(* IEC 61131-3 sources: machine-design-framework/examples/pick-glue-place/plc/generated, 2 files *)

(* ---- GVL_Cycle.st ---- *)
(* GENERATED from cycle.yaml - DO NOT EDIT. source-hash: bd31026db604f3bd *)
(* Commanded angles (deg). Effective timing = commanded + device delay; see GLUE-BEAD/PROD-* checks. *)
VAR_GLOBAL CONSTANT
    VACUUM_ON  : REAL := 10.0000;
    VACUUM_OFF : REAL := 222.0000;
    GLUE_GUN_ON  : REAL := 128.6400;
    GLUE_GUN_OFF : REAL := 130.4000;
    VAC_OK_CHECK : REAL := 26.0000;
    DOUBLE_SHEET_CHECK : REAL := 75.0000;
    HOST_BOOK_CHECK : REAL := 5.0000;
    HOST_SPINE_CHECK : REAL := 140.0000;
    BEAD_OK_CHECK : REAL := 148.0000;
    X_TRANSFER_OFFSET_MIN : REAL := 0.0000;   (* per-cycle offset range, mm *)
    X_TRANSFER_OFFSET_MAX : REAL := 15.0000;
    PARK_ANGLE : REAL := 355.0000;
END_VAR

(* ---- GVL_IO.st ---- *)
(* GENERATED from io_list.yaml - DO NOT EDIT. source-hash: db4df5e0d0977f7a *)
VAR_GLOBAL
    rAngle : REAL;   (* in  virtual *)
    rHostSpineOffset : REAL;   (* in  virtual *)
    rXOffset : REAL;   (* out  virtual *)
    xMasterRun : BOOL;   (* out  virtual *)
    xVacuum : BOOL;   (* out  DO1.0 EJECTOR *)
    xGlueGun : BOOL;   (* out  DO1.1 GLUE_VALVE *)
    xLampFault : BOOL;   (* out  DO1.2 LAMP_FAULT *)
    xVacOk : BOOL;   (* in  DI1.0 EJECTOR *)
    xDoubleSheet : BOOL;   (* in  DI1.1 DOUBLE_SENSOR *)
    xAirOk : BOOL;   (* in  DI1.2 AIR_SWITCH *)
    xGlueReady : BOOL;   (* in  DI1.3 GLUE_UNIT *)
    xBeadOk : BOOL;   (* in  DI1.7 BEAD_SENSOR *)
    xStartPb : BOOL;   (* in  DI1.4 OP_PANEL *)
    xStopPb : BOOL;   (* in  DI1.5 OP_PANEL *)
    xResetPb : BOOL;   (* in  DI1.6 OP_PANEL *)
    xHostBookPresent : BOOL;   (* in  DI2.0 BINDER_HANDSHAKE *)
    xGuardClosed : BOOL;   (* in  SDI1.0 GUARD_SWITCH *)
    xEStopOk : BOOL;   (* in  SDI1.1 ESTOP *)
END_VAR
